(* IEC 61131-3 sources: rusty/tests/lit/cfc/blocks/expression_input, 2 files *)

(* ---- main.st ---- *)
FUNCTION main : DINT
    expression_input();
    expression_input();
    // CHECK: a = 6, b = 20, sum = 26
    printf('a = %d, b = %d, sum = %d$N', expression_input.outA, expression_input.outB, expression_input.sum);
END_FUNCTION

(* ---- counter.st ---- *)
FUNCTION_BLOCK counter
VAR_INPUT
    step : DINT;
END_VAR
VAR_OUTPUT
    total : DINT;
END_VAR
    total := total + step;
END_FUNCTION_BLOCK
